FUNCTION_BLOCK XtsNctMover EXTENDS XtsMover IMPLEMENTS I_XtsNctMover
VAR
	_NctTask : XtsMoverNctTask;
	_NctTool : I_XtsNctTool;
END_VAR

(*FB_Init is always available implicitly and it is used primarily for initialization.
The return value is not evaluated. For a specific influence, you can also declare the
methods explicitly and provide additional code there with the standard initialization
code. You can evaluate the return value.*)
METHOD FB_Init : BOOL
VAR_INPUT
	(* TRUE: the retain variables are initialized (reset warm / reset cold)*)
	bInitRetains : BOOL;

	(* TRUE: the instance will be copied to the copy code afterward (online change)   *)
	bInCopyCode : BOOL;
	Name		: XtsCore.Core.T_MaxString;
	MoverData	: I_XtsMoverData;	  //Optional MoverData assignment
	System		: I_ContainXtsMovers; //Optional Self Registration with an Xts System
	NctTool		: I_XtsNctTool;		  //Optional Nct Tool assignment
END_VAR

VAR
	_Xts : I_XtsSystem;
END_VAR
IF __QUERYINTERFACE(System, _Xts) THEN
	_NctTask.XtsSystem := _Xts;
END_IF

_MoverTaskCollection.AddTask(_NctTask);

IF NctTool <> 0 THEN
	_NctTool := NctTool;	
	_NctTool.NctBaseUnit := _NctTask.Nct;
END_IF
END_METHOD

{attribute 'monitoring' := 'call'}
PROPERTY Nct : I_XtsNctBaseUnit
GET
Nct := _NctTask.Nct;
END_GET
SET
_NctTask.Nct := Nct;
END_SET
END_PROPERTY

{attribute 'monitoring' := 'call'}
PROPERTY NctReady : BOOL
GET
NctReady := _NctTask.NctReady;
END_GET
END_PROPERTY

PROPERTY NctTool : I_XtsNctTool
GET
NctTool := _NctTool;
END_GET
SET
_NctTool := NctTool;
END_SET
END_PROPERTY

END_FUNCTION_BLOCK

(* stored: Version 1.1.0.1, ProductVersion 3.1.4026.21
   POU XtsNctMover: Id {361a8abc-66b6-4b4e-9fdd-fc5a74404093}, SpecialFunc None
   Method FB_Init: Id {406517e2-0f46-4693-9585-eae7e9d931b1}
   Property Nct: Id {93ec728e-3bc4-4852-9ad1-1cdacb1d5f8e}
   Get Get: Id {cfada41e-e384-48dc-b94c-abdba5d22204}
   Set Set: Id {4e43e18c-5118-456e-ba33-99f90475346c}
   Property NctReady: Id {dfb3e380-7118-40e4-8d1c-f86d0c067bfb}
   Get Get: Id {ed933c79-3f10-4e97-8d12-2b31831f4660}
   Property NctTool: Id {10432d13-8be1-432b-9423-1ec35a1f27b3}
   Get Get: Id {7063d6f9-7703-4808-9a80-578d0e1da66d}
   Set Set: Id {0bc32cc0-9ffd-4927-aceb-51214750c5bf} *)
